PROGRAM MAIN
VAR
END_VAR


FunktionBlockDiagram();

END_PROGRAM

(* stored: Version 1.1.0.1
   POU MAIN: Id {339c9723-049f-4d8c-a8c3-4bc9c78b41ed}, SpecialFunc None *)
